Fanuc KAREL source: KT00236.KL

PROGRAM KT00236
%NOLOCKGROUP
VAR
  I1: INTEGER
  I2: INTEGER
  OUT: INTEGER
BEGIN
  I1 = 2
  I2 = 3
  I1 = 2
  I2 = 3
  OUT = I1 OR I2
END KT00236
